(* IEC 61131-3 sources: sis-interlock-demo/src/POUs/Sis/F_SisBit, 2 files *)

(* ---- F_SisBit.decl.st ---- *)
// Назначение: бит маски по индексу с единицы: бит uiIdx − 1; uiIdx вне 1..16 — FALSE.
// Автор:      kr0nsch
// Версия:     0.1.0
// Документ:   docs/DESIGN.md, раздел «8.2 Функции работы с битами»
// ВНИМАНИЕ:   код демонстрационный и не предназначен для систем безопасности. Реальная ПАЗ
//             требует определения SIL, сертифицированных аппаратных и программных средств
//             и валидации по ГОСТ Р МЭК 61511.
FUNCTION F_SisBit : BOOL
VAR_INPUT
    wMask : WORD;    // маска
    uiIdx : UINT;    // индекс причины или следствия, 1..16
END_VAR

(* ---- F_SisBit.impl.st ---- *)
IF uiIdx >= 1 AND uiIdx <= GVL_Const.WORD_BITS THEN
    F_SisBit := (wMask AND SHL(GVL_Const.WORD_BIT0, uiIdx - 1)) <> 0;
ELSE
    F_SisBit := FALSE;
END_IF
